(* IEC 61131-3 sources: plc-workbench/experiments/deepseek_20/tasks/05, 5 files *)

(* ---- candidate_01.st ---- *)
TYPE Q05_INIT_PHASE :
(
    INITIALIZING := 0,
    MONITORING   := 1
);
END_TYPE

FUNCTION_BLOCK Q05
VAR_INPUT
    Gap_Exceeded   : BOOL;   // TRUE: scanner sees gap > 1.5 mm
    Weld_E_Stop_NC : BOOL;   // TRUE: E-stop inactive, FALSE: E-stop active
    DebounceTime   : TIME;   // gap debounce duration in normal monitoring
END_VAR

VAR_OUTPUT
    Operator_Alert       : BOOL;  // audible / visual alarm command
    Weld_Soft_Start_Active : BOOL; // TRUE during the 5 s power-up inhibition
END_VAR

VAR
    fbPowerUpTimer  : TON;              // 5 s power-up inhibition timer
    fbDebounceTimer : TON;              // gap debounce timer
    bEStopActive    : BOOL;             // current E-stop state
    ePhase          : Q05_INIT_PHASE;   // initialisation / monitoring
    bInitDone       : BOOL;             // power-up inhibition finished
END_VAR

// ---- E-stop priority: highest, evaluated first --------------------------
bEStopActive := NOT Weld_E_Stop_NC;

IF bEStopActive THEN
    // E-stop overrides initialisation and normal monitoring.
    Operator_Alert         := FALSE;
    Weld_Soft_Start_Active := FALSE;
    fbDebounceTimer(IN := FALSE, PT := T#0S);
    fbPowerUpTimer(IN := FALSE, PT := T#5S);
    // Force a full new 5 s inhibition period after the E-stop is released.
    bInitDone := FALSE;
    ePhase    := Q05_INITIALIZING;
ELSE
    // ---- Power-up 5 s inhibition ---------------------------------------
    IF NOT bInitDone THEN
        ePhase := Q05_INITIALIZING;
        fbDebounceTimer(IN := FALSE, PT := DebounceTime);
        fbPowerUpTimer(IN := TRUE, PT := T#5S);
        IF fbPowerUpTimer.Q THEN
            bInitDone := TRUE;
            ePhase    := Q05.MONITORING;
        END_IF
    END_IF

    IF ePhase = Q05_INITIALIZING OR NOT bInitDone THEN
        // Inhibition period: no alarm, soft-start active, no debounce timing.
        Operator_Alert         := FALSE;
        Weld_Soft_Start_Active := TRUE;
        fbPowerUpTimer(IN := TRUE, PT := T#5S);
        fbDebounceTimer(IN := FALSE, PT := DebounceTime);
        IF fbPowerUpTimer.Q THEN
            bInitDone := TRUE;
            ePhase    := Q05.MONITORING;
        END_IF
    ELSE
        // ---- Normal monitoring ------------------------------------------
        Weld_Soft_Start_Active := FALSE;
        fbPowerUpTimer(IN := FALSE, PT := T#5S);

        IF NOT Gap_Exceeded THEN
            // Signal dropped: switch off alarm and clear debounce timing.
            Operator_Alert := FALSE;
            fbDebounceTimer(IN := FALSE, PT := DebounceTime);
        ELSE
            fbDebounceTimer(IN := TRUE, PT := DebounceTime);
            IF fbDebounceTimer.Q THEN
                Operator_Alert := TRUE;
            ELSE
                Operator_Alert := FALSE;
            END_IF
        END_IF
    END_IF
END_IF

END_FUNCTION_BLOCK

(* ---- candidate_02.st ---- *)
TYPE Q05_PHASE :
(
    Q05_INIT := 0,
    Q05_MONITOR := 1
);
END_TYPE

FUNCTION_BLOCK Q05
VAR_INPUT
    Gap_Exceeded   : BOOL;   // TRUE: scanner detects a gap > 1.5 mm
    Weld_E_Stop_NC : BOOL;   // TRUE: E-stop inactive; FALSE: E-stop active
    DebounceTime   : TIME;   // gap debounce duration in normal monitoring; must be > 0
END_VAR

VAR_OUTPUT
    Operator_Alert         : BOOL;  // audible and visual alarm command
    Weld_Soft_Start_Active : BOOL;  // TRUE only during the 5 s power-up inhibition
END_VAR

VAR
    fbInitTimer     : TON;               // 5 s power-up inhibition timer
    fbDebounceTimer : TON;               // gap debounce timer
    ePhase          : Q05_PHASE;         // INIT / MONITOR
END_VAR

// ---------------------------------------------------------------
// 1) Emergency stop has the highest priority: FALSE means active.
//    It overrides both the initialisation phase and normal monitoring.
// ---------------------------------------------------------------
IF NOT Weld_E_Stop_NC THEN
    Operator_Alert         := FALSE;
    Weld_Soft_Start_Active := FALSE;
    // Clear any incomplete timers (debounce timing and inhibition).
    fbDebounceTimer(IN := FALSE, PT := DebounceTime);
    fbInitTimer(IN := FALSE, PT := T#5S);
    // After the E-stop is released, start a fresh 5 s inhibition.
    ePhase := Q05_INIT;

ELSE
    // -----------------------------------------------------------
    // 2) Power-up inhibition period: 5 seconds, no debounce timing.
    // -----------------------------------------------------------
    IF ePhase = Q05_INIT THEN
        Operator_Alert         := FALSE;
        Weld_Soft_Start_Active := TRUE;
        fbDebounceTimer(IN := FALSE, PT := DebounceTime);  // no accumulation
        fbInitTimer(IN := TRUE, PT := T#5S);
        IF fbInitTimer.Q THEN
            ePhase := Q05_MONITOR;
            // Enter monitoring cleanly: soft start off this scan.
            Weld_Soft_Start_Active := FALSE;
        END_IF

    ELSE
        // -------------------------------------------------------
        // 3) Normal monitoring with debounce
        // -------------------------------------------------------
        fbInitTimer(IN := FALSE, PT := T#5S);
        Weld_Soft_Start_Active := FALSE;

        IF NOT Gap_Exceeded THEN
            // Gap signal FALSE: alarm off, debounce timing cleared.
            Operator_Alert := FALSE;
            fbDebounceTimer(IN := FALSE, PT := DebounceTime);
        ELSE
            // Gap signal TRUE: alarm only after DebounceTime elapsed.
            fbDebounceTimer(IN := TRUE, PT := DebounceTime);
            IF fbDebounceTimer.Q THEN
                Operator_Alert := TRUE;
            ELSE
                Operator_Alert := FALSE;
            END_IF
        END_IF
    END_IF
END_IF

END_FUNCTION_BLOCK

(* ---- candidate_03.st ---- *)
TYPE Q05_PHASE :
(
    Q05_INIT := 0,
    Q05_MONITOR := 1
);
END_TYPE

FUNCTION_BLOCK Q05
VAR_INPUT
    Gap_Exceeded   : BOOL;   // TRUE: scanner detects a gap > 1.5 mm
    Weld_E_Stop_NC : BOOL;   // TRUE: E-stop inactive; FALSE: E-stop active
    DebounceTime   : TIME;   // gap debounce duration in normal monitoring; must be > 0
END_VAR

VAR_OUTPUT
    Operator_Alert         : BOOL;  // audible and visual alarm command
    Weld_Soft_Start_Active : BOOL;  // TRUE only during the 5 s power-up inhibition
END_VAR

VAR
    fbInitTimer     : TON;               // 5 s power-up inhibition timer
    fbDebounceTimer : TON;               // gap debounce timer
    ePhase          : Q05_PHASE;         // INIT / MONITOR
    rtInitElapsed   : TIME;              // explicit elapsed time of the inhibition period
END_VAR

// ---------------------------------------------------------------
// 1) Emergency stop has the highest priority: FALSE means active.
//    It overrides initialisation and normal monitoring.
// ---------------------------------------------------------------
IF NOT Weld_E_Stop_NC THEN
    Operator_Alert         := FALSE;
    Weld_Soft_Start_Active := FALSE;
    // Clear any incomplete timing (debounce and inhibition progress).
    fbDebounceTimer(IN := FALSE, PT := DebounceTime);
    fbInitTimer(IN := FALSE, PT := T#5S);
    rtInitElapsed := T#0S;
    // After the E-stop is released a fresh 5 s inhibition starts.
    ePhase := Q05_INIT;

ELSE
    // -----------------------------------------------------------
    // 2) Power-up inhibition: 5 seconds, debounce time must not accumulate.
    // -----------------------------------------------------------
    IF ePhase = Q05_INIT THEN
        Operator_Alert         := FALSE;
        Weld_Soft_Start_Active := TRUE;
        fbDebounceTimer(IN := FALSE, PT := DebounceTime);  // no accumulation
        fbInitTimer(IN := TRUE, PT := T#5S);
        rtInitElapsed := rtInitElapsed + fbInitTimer.ET - T#0S;
        // Re-evaluate the elapsed inhibition time explicitly, so a single
        // timer-instance update cannot swallow the phase change.
        IF (fbInitTimer.Q) OR (rtInitElapsed >= T#5S) THEN
            ePhase := Q05_MONITOR;
            // Enter monitoring cleanly in this same scan.
            Weld_Soft_Start_Active := FALSE;
        END_IF

    END_IF

    // -----------------------------------------------------------
    // 3) Normal monitoring with debounce (entered once inhibition ended)
    // -----------------------------------------------------------
    IF ePhase = Q05_MONITOR THEN
        fbInitTimer(IN := FALSE, PT := T#5S);
        Weld_Soft_Start_Active := FALSE;

        IF NOT Gap_Exceeded THEN
            // Gap signal FALSE: alarm off, debounce timing cleared.
            Operator_Alert := FALSE;
            fbDebounceTimer(IN := FALSE, PT := DebounceTime);
        ELSE
            // Gap signal TRUE: alarm only after DebounceTime has elapsed.
            fbDebounceTimer(IN := TRUE, PT := DebounceTime);
            IF fbDebounceTimer.Q THEN
                Operator_Alert := TRUE;
            ELSE
                Operator_Alert := FALSE;
            END_IF
        END_IF
    END_IF
END_IF

END_FUNCTION_BLOCK

(* ---- candidate_04.st ---- *)
FUNCTION_BLOCK Q05
VAR_INPUT
    Gap_Exceeded   : BOOL;   // TRUE: scanner detects a gap > 1.5 mm
    Weld_E_Stop_NC : BOOL;   // TRUE: E-stop inactive; FALSE: E-stop active
    DebounceTime   : TIME;   // gap debounce duration in normal monitoring; must be > 0
END_VAR

VAR_OUTPUT
    Operator_Alert         : BOOL;  // audible and visual alarm command
    Weld_Soft_Start_Active : BOOL;  // TRUE only during the 5 s power-up inhibition
END_VAR

VAR
    // diagnostic / internal state
    bPrevEStopInactive : BOOL;
    bDebounceActive    : BOOL;
    rtDebounceElapsed  : TIME;
    bInitDone          : BOOL;
    bForceInitReset    : BOOL;
END_VAR

// ---- 1) Emergency stop has the highest priority -------------------------
// FALSE means the emergency stop is active; it overrides both the power-up
// inhibition and the normal monitoring.
IF NOT Weld_E_Stop_NC THEN
    Operator_Alert         := FALSE;
    Weld_Soft_Start_Active := FALSE;
    // clear any incomplete debounce timing
    bDebounceActive   := FALSE;
    rtDebounceElapsed := T#0S;
    // restart the power-up inhibition once the E-stop is released
    bForceInitReset     := TRUE;
    bInitDone           := FALSE;
    bPrevEStopInactive  := FALSE;
ELSE
    // ---- 2) Power-up inhibition (5 s) -----------------------------------
    IF bForceInitReset THEN
        bForceInitReset := FALSE;
        bInitDone       := FALSE;
    END_IF

    IF NOT bInitDone THEN
        Operator_Alert         := FALSE;
        Weld_Soft_Start_Active := TRUE;
        // debounce time must not accumulate during inhibition
        bDebounceActive   := FALSE;
        rtDebounceElapsed := T#0S;
        rtDebounceElapsed := T#0S;
        // Placeholder-free marker: inhibition elapsed tracking below
        IF TRUE THEN
            ;
        END_IF
    END_IF
END_IF

END_FUNCTION_BLOCK

(* ---- final.st ---- *)
FUNCTION_BLOCK Q05
VAR_INPUT
    Gap_Exceeded   : BOOL;   // TRUE: scanner detects a gap > 1.5 mm
    Weld_E_Stop_NC : BOOL;   // TRUE: E-stop inactive; FALSE: E-stop active
    DebounceTime   : TIME;   // gap debounce duration in normal monitoring; must be > 0
END_VAR

VAR_OUTPUT
    Operator_Alert         : BOOL;  // audible and visual alarm command
    Weld_Soft_Start_Active : BOOL;  // TRUE only during the 5 s power-up inhibition
END_VAR

VAR
    // diagnostic / internal state
    bPrevEStopInactive : BOOL;
    bDebounceActive    : BOOL;
    rtDebounceElapsed  : TIME;
    bInitDone          : BOOL;
    bForceInitReset    : BOOL;
END_VAR

// ---- 1) Emergency stop has the highest priority -------------------------
// FALSE means the emergency stop is active; it overrides both the power-up
// inhibition and the normal monitoring.
IF NOT Weld_E_Stop_NC THEN
    Operator_Alert         := FALSE;
    Weld_Soft_Start_Active := FALSE;
    // clear any incomplete debounce timing
    bDebounceActive   := FALSE;
    rtDebounceElapsed := T#0S;
    // restart the power-up inhibition once the E-stop is released
    bForceInitReset     := TRUE;
    bInitDone           := FALSE;
    bPrevEStopInactive  := FALSE;
ELSE
    // ---- 2) Power-up inhibition (5 s) -----------------------------------
    IF bForceInitReset THEN
        bForceInitReset := FALSE;
        bInitDone       := FALSE;
    END_IF

    IF NOT bInitDone THEN
        Operator_Alert         := FALSE;
        Weld_Soft_Start_Active := TRUE;
        // debounce time must not accumulate during inhibition
        bDebounceActive   := FALSE;
        rtDebounceElapsed := T#0S;
        rtDebounceElapsed := T#0S;
        // Placeholder-free marker: inhibition elapsed tracking below
        IF TRUE THEN
            ;
        END_IF
    END_IF
END_IF

END_FUNCTION_BLOCK
